Universal Robots URScript: T003_qwen2.5-coder_32b_baseline_rep1_retry2.urscript

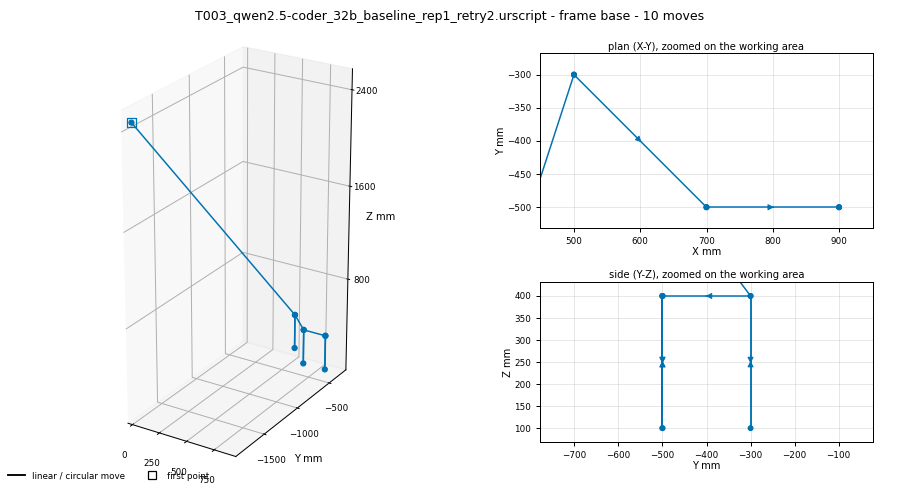
[picture p0: tool path of T003_qwen2.5-coder_32b_baseline_rep1_retry2.urscript in frame base, 10 of 10 moves have a stored position in this frame; points joined in program order, loops and branches not executed]
def task_eur_pallet()
    # Home position
    movej(p[0.000, -1.837, 2.459, 0.000, 2.618, 0.000], a=1.2, v=1.0)

    # Approach conveyor pick — above
    movel(p[0.500, -0.300, 0.400, 0.000, 2.618, 0.000], a=1.2, v=0.25)

    # Descend to pick
    movel(p[0.500, -0.300, 0.100, 0.000, 2.618, 0.000], a=1.2, v=0.1)

    # Lift from conveyor
    movel(p[0.500, -0.300, 0.400, 0.000, 2.618, 0.000], a=1.2, v=0.2)

    # Transit to pallet position (0,0)
    movel(p[0.700, -0.500, 0.400, 0.000, 2.618, 0.000], a=1.2, v=0.28)

    # Place on pallet (position 0,0)
    movel(p[0.700, -0.500, 0.100, 0.000, 2.618, 0.000], a=1.2, v=0.1)

    # Lift from pallet
    movel(p[0.700, -0.500, 0.400, 0.000, 2.618, 0.000], a=1.2, v=0.2)

    # Transit to next pallet position (1,0)
    movel(p[0.900, -0.500, 0.400, 0.000, 2.618, 0.000], a=1.2, v=0.28)

    # Place on pallet (position 1,0)
    movel(p[0.900, -0.500, 0.100, 0.000, 2.618, 0.000], a=1.2, v=0.1)

    # Lift from pallet
    movel(p[0.900, -0.500, 0.400, 0.000, 2.618, 0.000], a=1.2, v=0.2)
end

task_eur_pallet()
